{attribute 'qualified_only'}
VAR_GLOBAL
	nDrumsFilled : UDINT;
	bEStop AT %I* : BOOL;
END_VAR
VAR_GLOBAL CONSTANT
	MAX_MODULES : INT := 16;	// sizing constant: the runtime exports it without a READONLY flag
END_VAR

(* stored: Version 1.1.0.1, ProductVersion 3.1.4024.12
   GVL GVL_Machine: Id {aaaaaaaa-0000-0000-0000-000000000009} *)
